Fanuc KAREL source: kt00120.KL

-- PROVISIONAL review KL for V1013-1; original PC SHA256 2310a2459e2e624cebf9babd90a57d4f4b8312a8a4986142b0a6b1c859b8aaad
-- Incomplete behavior may be omitted. Consult companion uncertainty JSON. Do not deploy.
PROGRAM KT00120
%NOLOCKGROUP
VAR
  OUT : REAL
-- UNRESOLVED_DECL Y1 type=002018
-- UNRESOLVED_DECL H2 type=002017
BEGIN
  -- UNRESOLVED_PC offsets 5-19; opcodes 2E,22,9D,33,B2
  -- UNRESOLVED_PC offsets 24-38; opcodes 2E,22,9D,33,B4
  -- UNRESOLVED_PC offsets 43-72; opcodes 22,9D,33,B1,22,9D,33,B3,64,29,64,29,6C,23
  -- UNRESOLVED_PC offsets 77-81; opcodes 7F
END KT00120
